// TIA Portal V19 export
VAR_GLOBAL   // PLC tag table "IO_Tags"
   "ZSO-112B" AT %I100.2 : Bool;   // Válvula entrada de meladura cruda - Confirmación Apertura
   "ZSO-112A" AT %I100.3 : Bool;   // Válvula entrada de meladura clarificada - Confirmación Apertura
   "ZSO-105" AT %I100.4 : Bool;   // Válvula entrada de semilla - Confirmación Apertura
   "ZSO-103" AT %I100.5 : Bool;   // Válvula rompevacío - Confirmación Apertura
   "ZSO-109" AT %I100.6 : Bool;   // Válvula de descarga - Confirmación Apertura
   "ZSO-104" AT %I100.7 : Bool;   // Vávula inyección de colada - Confirmación Apertura
   "ZSO-108" AT %I101.0 : Bool;   // Válvula corte tacho 3 al 2 - Confirmación Apertura
   "YI-101" AT %I101.1 : Bool;   // Agitador - Confirmación de run
   "YT-101" AT %I101.2 : Bool;   // Agitador - Disparo
   "ZSO-102" AT %I101.5 : Bool;   // Válvula soplo - Confirmación Apertura
   "TSV-102" AT %Q100.5 : Bool;   // Válvula soplo - Comando Apertura/Cierre
   "XSV-112B" AT %Q100.6 : Bool;   // Válvula entrada de meladura cruda - Comando Apertura/Cierre
   "XSV-112A" AT %Q100.7 : Bool;   // Válvula entrada de meladura clarificada - Comando Apertura/Cierre
   "XSV-105" AT %Q101.0 : Bool;   // Válvula entrada de semilla - Comando Apertura/Cierre
   "PSV-103" AT %Q101.1 : Bool;   // Válvula rompevacío - Comando Apertura/Cierre
   "LSV-109" AT %Q101.2 : Bool;   // Válvula de descarga - Comando Apertura/Cierre
   "XSV-104" AT %Q101.3 : Bool;   // Vávula inyección de colada - Comando Apertura/Cierre
   "XSV-108" AT %Q101.4 : Bool;   // Válvula corte tacho 3 al 2 - Comando Apertura/Cierre
   "M-101" AT %Q101.5 : Bool;   // Agitador - Comando Start/Stop
   "LT-112" AT %IW256 : Int;   // Nivel Tacho - Lectura
   "PT-110" AT %IW258 : Int;   // Presión de vacío - Lectura
   "PT-113" AT %IW260 : Int;   // Presion de vapor a calandria - Lectura
   "TT-114" AT %IW262 : Int;   // Temperatura del cuerpo - Lectura
   "TT-115" AT %IW264 : Int;   // Temperatura calandria - Lectura
   "AT-112" AT %IW266 : Int;   // Brix masa cocida - sonda microondas - Lectura
   "LCV-212" AT %QW256 : Int;   // Válvula entrada de meladura - Consigna análoga de apertura
   "DCV-211" AT %QW258 : Int;   // Válvula entrada vapor calandria - Consigna análoga de apertura
   "XCV-107" AT %QW260 : Int;   // Válvula entrada de agua caliente - Consigna análoga de apertura
   "PCV-210" AT %QW262 : Int;   // Válvula entrada de agua al condensador - Consigna análoga de apertura
   Tacho1_SM_Input AT %I0.0 : "Pan_From_SM";
   Tacho1_SM_Output AT %Q0.0 : "Pan_To_SM";
   Tacho2_SM_Input AT %I69.0 : "Pan_From_SM";
   Tacho2_SM_Output AT %Q41.0 : "Pan_To_SM";
   "ZSO-113" AT %I101.6 : Bool;   // Válvula de desagüe (futura)
   "XSV-113" AT %Q101.6 : Bool;   // Válvula de desagüe (futura)
   "LT-116" AT %IW268 : Int;   // Nivel recibidor de masa - Lectura
   "AT-112x" AT %IW270 : Int;   // Brix masa cocida - sonda microondas - Raw
   "YI-102" AT %I101.3 : Bool;   // Bomba vacío - Confirmación de run
   "M-102" AT %Q101.7 : Bool;   // Bomba vacío - Comando Start/Stop
   "YSH-000" AT %Q100.0 : Bool;   // Alarma visual
   "XSV-114" AT %Q100.3 : Bool;   // Valvula lavado sensores de brix
   "YSL-000" AT %Q100.1 : Bool;   // Advertencia visual
END_VAR
